Yaskawa INFORM job: -DEFRO-70_PRZYLACZE_60_STARE.JBI

/JOB
//NAME -DEFRO-70_PRZYLACZE_60_STARE
//POS
///NPOS 165,165,165,0,0,0
///TOOL 0
///POSTYPE PULSE
///PULSE
C00000=-281,-101163,-84214,3730,-80188,-1936
C00001=-283,-101162,-84213,3710,-80188,-1936
C00002=115939,-17843,-44700,-6904,-63515,59085
C00003=117854,12047,-44285,-6364,-54274,83125
C00004=118072,11991,-44277,-6360,-54292,83048
C00005=124625,19348,-37580,2226,-58698,65873
C00006=128138,4548,-53928,8815,-39472,48638
C00007=140958,30570,-37086,38951,-57450,21007
C00008=144303,30296,-42198,53003,-55772,9063
C00009=140286,42517,-25172,35381,-64941,20617
C00010=134888,48773,-14255,24473,-68176,15010
C00011=126216,57142,-1405,12520,-73831,-5965
C00012=119431,58070,-113,1607,-75333,-12308
C00013=112362,60124,-1581,-7248,-81906,-32507
C00014=102321,53890,-14377,-28322,-78386,-34401
C00015=102712,42577,-23807,-28139,-73777,-45229
C00016=111795,28445,-30470,-11492,-65646,-58750
C00017=113823,16078,-41175,-14074,-58178,-74794
C00018=114023,15964,-41317,-14088,-58122,-74856
C00019=114170,-2374,-36949,-11645,-74681,-76938
C00020=113314,-7643,-38017,-11019,-76954,88145
C00021=103795,24169,-32802,-5113,-62316,87115
C00022=105717,22963,-33847,-2915,-61383,82248
C00023=105949,12675,-44086,-6804,-51663,75716
C00024=112305,4286,-54083,4280,-38458,55374
C00025=119011,7063,-54209,24198,-38298,40510
C00026=126176,29519,-37310,40709,-52379,12824
C00027=124287,36853,-27992,32882,-57796,17661
C00028=118323,57808,-3223,17808,-73635,15605
C00029=113918,55938,-2510,14235,-71141,-2239
C00030=100452,57135,-1831,-9316,-72769,-11707
C00031=101122,66320,5615,-3405,-83775,-29323
C00032=90969,64062,-2652,-23907,-83052,-31977
C00033=91048,41774,-22566,-24453,-68601,-40164
C00034=95890,27642,-32117,-16170,-61880,-54638
C00035=99625,19836,-37924,-13704,-58629,-70011
C00036=99745,19765,-37997,-13694,-58605,-70048
C00037=99303,8604,-31154,-10952,-72489,-71699
C00038=89422,16015,-23794,-2157,-75183,91094
C00039=91342,36521,-20369,-2557,-66713,90648
C00040=96608,27573,-29625,3606,-58513,75053
C00041=104075,24092,-36197,17400,-51418,55933
C00042=113942,24510,-45627,50308,-45587,24643
C00043=113180,34271,-33600,43117,-51129,17495
C00044=105987,58297,-1625,19620,-69218,16598
C00045=102657,59844,2089,16796,-69099,938
C00046=91593,70320,13088,-1311,-78194,-10490
C00047=88532,80640,21579,-3911,-88822,-24498
C00048=80672,78287,14638,-19772,-88445,-29832
C00049=78449,68959,3821,-24282,-82660,-32911
C00050=77699,46922,-17540,-28065,-68732,-40538
C00051=80754,29721,-31897,-24408,-56253,-47712
C00052=85616,26363,-32270,-14653,-55936,-57384
C00053=85063,22114,-18753,-9149,-74798,-67250
C00054=72786,31521,-9549,-9445,-75352,93043
C00055=79344,46650,-9742,-3090,-64918,94922
C00056=79851,45963,-10489,-3142,-64795,94764
C00057=83555,34866,-22970,1140,-53515,77559
C00058=88637,21070,-41506,13142,-33787,59480
C00059=92546,17739,-49130,33624,-25291,42497
C00060=100296,32921,-36962,50214,-42105,29169
C00061=99518,40044,-26222,41163,-46688,21660
C00062=98807,50157,-13852,39808,-52940,6845
C00063=91319,71721,15887,17155,-70404,4779
C00064=77791,87178,32687,-9256,-82589,-4510
C00065=78950,98816,44020,-1274,-94156,-21475
C00066=71782,98188,39845,-16228,-95193,-28058
C00067=67733,74026,11935,-24954,-78838,-32081
C00068=70123,56840,-3457,-20485,-67729,-42469
C00069=71488,56179,-3109,-17368,-68202,-45369
C00070=72709,50202,-8538,-17621,-67542,-57502
C00071=75039,37514,-3449,-7701,-77257,-64173
C00072=74616,28156,-12897,-9694,-74827,92488
C00073=75521,47327,-9742,-11513,-65249,93468
C00074=83421,34104,-23568,1133,-53536,80045
C00075=88561,20457,-41927,13093,-33823,59529
C00076=92662,18115,-48904,33764,-25272,42413
C00077=97937,26210,-42655,47625,-35211,32454
C00078=99376,40032,-26365,41218,-46566,21666
C00079=100200,49079,-17087,46041,-52311,4065
C00080=91093,71344,15665,17037,-69989,4842
C00081=77993,87860,33884,-9296,-82933,-4594
C00082=79105,99458,45109,-1336,-94484,-21522
C00083=71734,96974,38291,-16203,-94882,-27999
C00084=67577,72994,10856,-25287,-78095,-32283
C00085=72681,51483,-6944,-14654,-65784,-51471
C00086=76109,49503,-7560,-9343,-66865,-57435
C00087=74844,35432,-1015,-7610,-79822,-64270
C00088=74616,28156,-12897,-9694,-74827,92488
C00089=90411,-2677,-20047,-11125,-84138,86440
C00090=90413,-2674,-20051,-11105,-84138,86441
C00091=137757,-12075,-30464,2646,-72394,74401
C00092=139263,-65150,-85436,14259,-28990,73053
C00093=136879,-25803,-69250,35998,-11820,63023
C00094=139290,-23505,-65815,37849,-15870,40588
C00095=138255,-25667,-68923,45072,-10125,18948
C00096=137540,-11621,-49291,15825,-29065,282
C00097=134494,-8817,-45605,4069,-31945,-3289
C00098=134604,-8591,-45393,4272,-32069,-3452
C00099=128608,-126,-37091,-12913,-41572,-17604
C00100=135365,-22598,-63276,22384,-16411,-55250
C00101=133643,-21758,-61840,7774,-18256,-58833
C00102=132849,-22230,-62300,-146,-18489,-67744
C00103=134650,-26769,-71812,22381,-6082,-94556
C00104=132637,-74135,-100376,4983,-10333,-85647
C00105=119687,-78067,-87939,-2788,-20735,84624
C00106=119992,-27745,-68017,-3051,-15116,84333
C00107=119030,-28696,-69591,-21999,-13157,75803
C00108=119146,-27568,-67331,-20983,-14326,49763
C00109=119106,-25320,-64288,-16073,-16150,28459
C00110=116990,-27787,-67992,-36968,-13306,28443
C00111=114451,-20387,-59191,-34974,-24024,21051
C00112=114289,-23226,-63137,-42813,-20195,20855
C00113=115755,-27101,-67787,-45506,-13897,17108
C00114=116631,-28534,-69574,-43897,-10967,13052
C00115=119721,-30747,-72526,-5019,-4908,-12317
C00116=124673,-29524,-70968,54153,-12690,-50315
C00117=110381,-14519,-53439,-34713,-36084,-50985
C00118=115065,-20808,-58231,-19385,-28009,-64203
C00119=113126,-78683,-102705,-45607,-16425,-60367
C00120=120908,-77676,-80309,7462,-22023,84016
C00121=119355,-30092,-72700,-7480,-8883,86833
C00122=119330,-30666,-73900,-37441,-7256,75668
C00123=119392,-31005,-74194,-36731,-7285,75171
C00124=119107,-25533,-64139,-15884,-16345,28370
C00125=118189,-11113,-47154,-8478,-33276,7215
C00126=118285,-13415,-49709,-5227,-31034,-7778
C00127=112204,-14619,-53166,-28572,-30616,-12922
C00128=112459,-20642,-60567,-34495,-24493,-27463
C00129=113253,-23242,-63602,-34662,-21946,-37788
C00130=117822,-27208,-67860,-16762,-15410,-62087
C00131=114088,-29625,-74008,-62760,-13130,-51071
C00132=113074,-79856,-103225,-44998,-16651,-60643
C00133=120443,-70015,-86553,-1670,-18639,84017
C00134=119855,-29453,-70963,-4444,-11447,85360
C00135=119350,-27114,-66909,-10824,-16764,76179
C00136=120538,-28712,-69581,-9042,-12118,60389
C00137=121453,-23804,-62042,-1822,-20367,42740
C00138=119104,-25714,-64462,-15988,-16245,28420
C00139=118127,-25090,-63854,-17709,-16479,10287
C00140=118054,-20647,-58029,-8598,-22594,-6818
C00141=116391,-17852,-55102,-12391,-26715,-16410
C00142=113676,-17333,-55635,-24105,-28107,-26621
C00143=114148,-20487,-59353,-25400,-25301,-39443
C00144=114654,-26064,-67349,-36235,-17702,-47147
C00145=115014,-30497,-76060,-73901,-10838,-47744
C00146=112648,-89264,-107216,-40476,-18619,-62704
C00147=115490,-77010,-93554,-11224,-18305,89052
C00148=125433,-24819,-64014,25600,-22035,67229
C00149=124409,-21324,-58576,14136,-26697,62401
C00150=126029,-28427,-71429,47699,-12406,35561
C00151=126376,-14543,-51553,17453,-33391,37954
C00152=119104,-25707,-64456,-15987,-16243,28419
C00153=102227,-21803,-62565,-47260,-20333,28942
C00154=103256,-22698,-63333,-30550,-15064,8897
C00155=100032,-11798,-50575,-26640,-29993,-6479
C00156=97406,-10335,-50320,-35130,-33056,-18084
C00157=102127,-19671,-59474,-25169,-24074,-49644
C00158=96594,-22492,-70681,-79494,-21703,-41695
C00159=112538,-91654,-108181,-39431,-19159,-63177
C00160=113545,-73371,-70378,-16072,-42358,69017
C00161=89593,-90202,-78264,-12204,-55560,23671
C00162=60247,-88344,-77535,-12630,-64499,59028
C00163=11932,-100155,-87763,417,-74819,10359
C00164=-281,-101163,-84214,3730,-80188,-1936
BC00000=570125
BC00001=868704
BC00002=878894
BC00003=878037
BC00004=878037
BC00005=878038
BC00006=878037
BC00007=878038
BC00008=878038
BC00009=878038
BC00010=878038
BC00011=878038
BC00012=878038
BC00013=878037
BC00014=878037
BC00015=878037
BC00016=878037
BC00017=878037
BC00018=878037
BC00019=878037
BC00020=912823
BC00021=878035
BC00022=878036
BC00023=878036
BC00024=878037
BC00025=878037
BC00026=878037
BC00027=878037
BC00028=878038
BC00029=878038
BC00030=878037
BC00031=878037
BC00032=878037
BC00033=878037
BC00034=878037
BC00035=878037
BC00036=878037
BC00037=878037
BC00038=878035
BC00039=878036
BC00040=878037
BC00041=878037
BC00042=878038
BC00043=878038
BC00044=878038
BC00045=878038
BC00046=878037
BC00047=878037
BC00048=878037
BC00049=878037
BC00050=878037
BC00051=878037
BC00052=878037
BC00053=878037
BC00054=878037
BC00055=878035
BC00056=878035
BC00057=877203
BC00058=877947
BC00059=878201
BC00060=878342
BC00061=878784
BC00062=877961
BC00063=877604
BC00064=878504
BC00065=878840
BC00066=878535
BC00067=877975
BC00068=879348
BC00069=879174
BC00070=879174
BC00071=878037
BC00072=915550
BC00073=913919
BC00074=916409
BC00075=916569
BC00076=916479
BC00077=916387
BC00078=916586
BC00079=915550
BC00080=915870
BC00081=916359
BC00082=916889
BC00083=917058
BC00084=916344
BC00085=916664
BC00086=916387
BC00087=915811
BC00088=915550
BC00089=915550
BC00090=915550
BC00091=915550
BC00092=915550
BC00093=915550
BC00094=915550
BC00095=915550
BC00096=915550
BC00097=915550
BC00098=915550
BC00099=915550
BC00100=915550
BC00101=915550
BC00102=915550
BC00103=915550
BC00104=915550
BC00105=915550
BC00106=915551
BC00107=915550
BC00108=915550
BC00109=915550
BC00110=915550
BC00111=915550
BC00112=915550
BC00113=915550
BC00114=915550
BC00115=915550
BC00116=915550
BC00117=915550
BC00118=915550
BC00119=915550
BC00120=954211
BC00121=953187
BC00122=954162
BC00123=954160
BC00124=954071
BC00125=953684
BC00126=953455
BC00127=953244
BC00128=953665
BC00129=953702
BC00130=953799
BC00131=953749
BC00132=953683
BC00133=992214
BC00134=992214
BC00135=992103
BC00136=991968
BC00137=992423
BC00138=992186
BC00139=992082
BC00140=991590
BC00141=991168
BC00142=991569
BC00143=992150
BC00144=992735
BC00145=991845
BC00146=991844
BC00147=1026906
BC00148=1030289
BC00149=1030277
BC00150=1030261
BC00151=1030281
BC00152=1030485
BC00153=997557
BC00154=991657
BC00155=991168
BC00156=991569
BC00157=992735
BC00158=991845
BC00159=1030552
BC00160=1030552
BC00161=1015004
BC00162=995119
BC00163=847363
BC00164=570125
EC00000=1163,0
EC00001=1166,0
EC00002=-1742,0
EC00003=-1741,0
EC00004=-1741,0
EC00005=-1743,0
EC00006=-1742,0
EC00007=-1741,0
EC00008=-1741,0
EC00009=-1741,0
EC00010=-1741,0
EC00011=-1741,0
EC00012=-1741,0
EC00013=-1741,0
EC00014=-1742,0
EC00015=-1742,0
EC00016=-1742,0
EC00017=-1741,0
EC00018=-1741,0
EC00019=-1741,0
EC00020=-1741,0
EC00021=-1745,0
EC00022=-1744,0
EC00023=-1743,0
EC00024=-1742,0
EC00025=-1742,0
EC00026=-1741,0
EC00027=-1741,0
EC00028=-1741,0
EC00029=-1741,0
EC00030=-1741,0
EC00031=-1741,0
EC00032=-1742,0
EC00033=-1742,0
EC00034=-1741,0
EC00035=-1741,0
EC00036=-1741,0
EC00037=-1741,0
EC00038=-1743,0
EC00039=-1742,0
EC00040=-1742,0
EC00041=-1742,0
EC00042=-1741,0
EC00043=-1741,0
EC00044=-1595,0
EC00045=-1742,0
EC00046=-1741,0
EC00047=-1741,0
EC00048=-1742,0
EC00049=-1742,0
EC00050=-1742,0
EC00051=-1742,0
EC00052=-1742,0
EC00053=-1741,0
EC00054=-1741,0
EC00055=-1743,0
EC00056=-1743,0
EC00057=-1742,0
EC00058=-1743,0
EC00059=-1742,0
EC00060=-1741,0
EC00061=-1741,0
EC00062=-1742,0
EC00063=-1742,0
EC00064=-1742,0
EC00065=-1741,0
EC00066=-1741,0
EC00067=-1741,0
EC00068=-1741,0
EC00069=-1741,0
EC00070=-1741,0
EC00071=-1741,0
EC00072=-1741,0
EC00073=-1742,0
EC00074=-1742,0
EC00075=-1743,0
EC00076=-1742,0
EC00077=-1741,0
EC00078=-1740,0
EC00079=-1742,0
EC00080=-1742,0
EC00081=-1742,0
EC00082=-1741,0
EC00083=-1741,0
EC00084=-1741,0
EC00085=-1742,0
EC00086=-1742,0
EC00087=-1741,0
EC00088=-1741,0
EC00089=-1741,0
EC00090=-84878,0
EC00091=-84879,0
EC00092=-84877,0
EC00093=-84877,0
EC00094=-84877,0
EC00095=-84877,0
EC00096=-84877,0
EC00097=-84877,0
EC00098=-84877,0
EC00099=-84877,0
EC00100=-84877,0
EC00101=-84877,0
EC00102=-84877,0
EC00103=-84877,0
EC00104=-84877,0
EC00105=-84877,0
EC00106=-84878,0
EC00107=-84877,0
EC00108=-84877,0
EC00109=-84877,0
EC00110=-84877,0
EC00111=-84877,0
EC00112=-84877,0
EC00113=-84877,0
EC00114=-84877,0
EC00115=-84877,0
EC00116=-84877,0
EC00117=-84877,0
EC00118=-84877,0
EC00119=-84877,0
EC00120=-84877,0
EC00121=-84878,0
EC00122=-84877,0
EC00123=-84877,0
EC00124=-84877,0
EC00125=-84877,0
EC00126=-84877,0
EC00127=-84877,0
EC00128=-84877,0
EC00129=-84877,0
EC00130=-84877,0
EC00131=-84877,0
EC00132=-84877,0
EC00133=-84877,0
EC00134=-84877,0
EC00135=-84877,0
EC00136=-84877,0
EC00137=-84877,0
EC00138=-84877,0
EC00139=-84877,0
EC00140=-84877,0
EC00141=-84877,0
EC00142=-84877,0
EC00143=-84877,0
EC00144=-84877,0
EC00145=-84877,0
EC00146=-84877,0
EC00147=-84877,0
EC00148=-84877,0
EC00149=-84877,0
EC00150=-84877,0
EC00151=-84877,0
EC00152=-84877,0
EC00153=-84877,0
EC00154=-84877,0
EC00155=-84877,0
EC00156=-84877,0
EC00157=-84877,0
EC00158=-84877,0
EC00159=-84877,0
EC00160=-84877,0
EC00161=-1879,0
EC00162=-1342,0
EC00163=498,0
EC00164=1163,0
//INST
///DATE 2025/05/12 13:13
///COMM OZZ
///ATTR SC,RW
///GROUP1 RB1,BS1
///GROUP2 ST1
NOP
MOVJ C00000 BC00000 VJ=70.00 DEC=20  +MOVJ EC00000 VJ=70.00
MOVJ C00001 BC00001 VJ=40.00 DEC=20  +MOVJ EC00001 VJ=40.00
MOVJ C00002 BC00002 VJ=70.00 DEC=20  +MOVJ EC00002 VJ=70.00
MOVJ C00003 BC00003 VJ=40.00 DEC=20  +MOVJ EC00003 VJ=70.00
MACRO1 MJ#(0) ARGF8
WVON WEV#(1)
ARCON
MOVC C00004 BC00004 V=4.2 DEC=20  +MOVJ EC00004 VJ=70.00
MOVC C00005 BC00005 V=4.2 DEC=20  +MOVJ EC00005 VJ=30.00
MOVC C00006 BC00006 V=4.2 DEC=20  +MOVJ EC00006 VJ=30.00
MOVC C00007 BC00007 V=4.2 DEC=20  +MOVJ EC00007 VJ=30.00
MOVC C00008 BC00008 V=4.2 DEC=20  +MOVJ EC00008 VJ=30.00
MOVC C00009 BC00009 V=4.2 DEC=20  +MOVJ EC00009 VJ=0.78
MOVC C00010 BC00010 V=4.2 DEC=20  +MOVJ EC00010 VJ=30.00
MOVC C00011 BC00011 V=4.2 DEC=20  +MOVJ EC00011 VJ=30.00
MOVC C00012 BC00012 V=4.2 DEC=20  +MOVJ EC00012 VJ=30.00
MOVC C00013 BC00013 V=4.2 DEC=20  +MOVJ EC00013 VJ=30.00
MOVC C00014 BC00014 V=4.2 DEC=20  +MOVJ EC00014 VJ=30.00
MOVC C00015 BC00015 V=4.2 DEC=20  +MOVJ EC00015 VJ=30.00
MOVC C00016 BC00016 V=4.2 DEC=20  +MOVJ EC00016 VJ=30.00
MOVC C00017 BC00017 V=4.2 DEC=20  +MOVJ EC00017 VJ=30.00
MOVJ C00018 BC00018 VJ=30.00 DEC=20  +MOVJ EC00018 VJ=30.00
WVOF
ARCOF
MOVJ C00019 BC00019 VJ=40.00 DEC=20  +MOVJ EC00019 VJ=40.00
MOVJ C00020 BC00020 VJ=70.00 DEC=20  +MOVJ EC00020 VJ=0.78
MOVJ C00021 BC00021 VJ=30.00 DEC=20  +MOVJ EC00021 VJ=0.78
MACRO1 MJ#(0) ARGF8
WVON WEV#(1)
ARCON
MOVC C00022 BC00022 V=4.2 DEC=20  +MOVJ EC00022 VJ=0.78
MOVC C00023 BC00023 V=4.2 DEC=20  +MOVJ EC00023 VJ=0.78
MOVC C00024 BC00024 V=4.2 DEC=20  +MOVJ EC00024 VJ=30.00
MOVC C00025 BC00025 V=4.2 DEC=20  +MOVJ EC00025 VJ=30.00
MOVC C00026 BC00026 V=5.0 DEC=20  +MOVJ EC00026 VJ=30.00
MOVC C00027 BC00027 V=4.2 DEC=20  +MOVJ EC00027 VJ=0.78
MOVC C00028 BC00028 V=4.2 DEC=20  +MOVJ EC00028 VJ=30.00
MOVC C00029 BC00029 V=4.2 DEC=20  +MOVJ EC00029 VJ=30.00
MOVC C00030 BC00030 V=4.2 DEC=20  +MOVJ EC00030 VJ=30.00
MOVC C00031 BC00031 V=4.2 DEC=20  +MOVJ EC00031 VJ=30.00
MOVC C00032 BC00032 V=4.2 DEC=20  +MOVJ EC00032 VJ=30.00
MOVC C00033 BC00033 V=4.2 DEC=20  +MOVJ EC00033 VJ=30.00
MOVC C00034 BC00034 V=4.2 DEC=20  +MOVJ EC00034 VJ=30.00
MOVC C00035 BC00035 V=4.2 DEC=20  +MOVJ EC00035 VJ=30.00
MOVJ C00036 BC00036 VJ=25.00 DEC=20  +MOVJ EC00036 VJ=30.00
WVOF
ARCOF
MOVJ C00037 BC00037 VJ=30.00 DEC=20  +MOVJ EC00037 VJ=30.00
MOVJ C00038 BC00038 VJ=30.00 DEC=20  +MOVJ EC00038 VJ=30.00
MOVJ C00039 BC00039 VJ=30.00 DEC=20  +MOVJ EC00039 VJ=30.00
WVON WEV#(1)
ARCON
MOVC C00040 BC00040 V=4.2 DEC=20  +MOVJ EC00040 VJ=30.00
MOVC C00041 BC00041 V=4.2 DEC=20  +MOVJ EC00041 VJ=30.00
MOVC C00042 BC00042 V=4.2 DEC=20  +MOVJ EC00042 VJ=30.00
MOVC C00043 BC00043 V=4.2 DEC=20  +MOVJ EC00043 VJ=30.00
MOVC C00044 BC00044 V=4.2 DEC=20  +MOVJ EC00044 VJ=30.00
MOVC C00045 BC00045 V=4.2 DEC=20  +MOVJ EC00045 VJ=30.00
MOVC C00046 BC00046 V=4.2 DEC=20  +MOVJ EC00046 VJ=30.00
MOVC C00047 BC00047 V=4.2 DEC=20  +MOVJ EC00047 VJ=30.00
MOVC C00048 BC00048 V=4.2 DEC=20  +MOVJ EC00048 VJ=30.00
MOVC C00049 BC00049 V=4.2 DEC=20  +MOVJ EC00049 VJ=0.78
MOVC C00050 BC00050 V=5.8 DEC=20  +MOVJ EC00050 VJ=30.00
MOVC C00051 BC00051 V=4.2 DEC=20  +MOVJ EC00051 VJ=0.78
MOVC C00052 BC00052 V=4.2 DEC=20  +MOVJ EC00052 VJ=30.00
ARCOF
WVOF
MOVJ C00053 BC00053 VJ=30.00 DEC=20  +MOVJ EC00053 VJ=30.00
MOVJ C00054 BC00054 VJ=30.00 DEC=20  +MOVJ EC00054 VJ=30.00
MOVJ C00055 BC00055 VJ=30.00 DEC=20  +MOVJ EC00055 VJ=30.00
WVON WEV#(1)
ARCON
MOVC C00056 BC00056 V=4.2 DEC=20  +MOVJ EC00056 VJ=0.78
MOVC C00057 BC00057 V=4.2 DEC=20  +MOVJ EC00057 VJ=0.78
MOVC C00058 BC00058 V=4.2 DEC=20  +MOVJ EC00058 VJ=0.78
MOVC C00059 BC00059 V=4.2 DEC=20  +MOVJ EC00059 VJ=0.78
MOVC C00060 BC00060 V=4.2 DEC=20  +MOVJ EC00060 VJ=0.78
MOVC C00061 BC00061 V=4.2 DEC=20  +MOVJ EC00061 VJ=0.78
MOVC C00062 BC00062 V=4.2 DEC=20  +MOVJ EC00062 VJ=0.78
MOVC C00063 BC00063 V=4.2 DEC=20  +MOVJ EC00063 VJ=0.78
MOVC C00064 BC00064 V=4.2 DEC=20  +MOVJ EC00064 VJ=0.78
MOVC C00065 BC00065 V=4.2 DEC=20  +MOVJ EC00065 VJ=0.78
MOVC C00066 BC00066 V=4.2 DEC=20  +MOVJ EC00066 VJ=0.78
MOVC C00067 BC00067 V=4.2 DEC=20  +MOVJ EC00067 VJ=0.78
MOVC C00068 BC00068 V=4.2 DEC=20  +MOVJ EC00068 VJ=0.78
MOVC C00069 BC00069 V=4.2 DEC=20  +MOVJ EC00069 VJ=0.78
MOVC C00070 BC00070 V=4.2 DEC=20  +MOVJ EC00070 VJ=0.78
WVOF
ARCOF
MOVJ C00071 BC00071 VJ=30.00 DEC=20  +MOVJ EC00071 VJ=30.00
MOVJ C00072 BC00072 VJ=30.00 DEC=20  +MOVJ EC00072 VJ=30.00
MOVJ C00073 BC00073 VJ=30.00 DEC=20  +MOVJ EC00073 VJ=30.00
WVON WEV#(1)
ARCON
MOVC C00074 BC00074 V=4.2 DEC=20  +MOVJ EC00074 VJ=30.00
MOVC C00075 BC00075 V=4.2 DEC=20  +MOVJ EC00075 VJ=30.00
MOVC C00076 BC00076 V=4.2 DEC=20  +MOVJ EC00076 VJ=40.00
MOVC C00077 BC00077 V=4.2 DEC=20  +MOVJ EC00077 VJ=30.00
MOVC C00078 BC00078 V=4.2 DEC=20  +MOVJ EC00078 VJ=25.00
MOVC C00079 BC00079 V=4.2 DEC=20  +MOVJ EC00079 VJ=30.00
MOVC C00080 BC00080 V=4.2 DEC=20  +MOVJ EC00080 VJ=70.00
MOVC C00081 BC00081 V=4.2 DEC=20  +MOVJ EC00081 VJ=30.00
MOVC C00082 BC00082 V=4.2 DEC=20  +MOVJ EC00082 VJ=30.00
MOVC C00083 BC00083 V=4.2 DEC=20  +MOVJ EC00083 VJ=30.00
MOVC C00084 BC00084 V=4.2 DEC=20  +MOVJ EC00084 VJ=30.00
MOVC C00085 BC00085 V=4.2 DEC=20  +MOVJ EC00085 VJ=0.78
MOVC C00086 BC00086 V=4.2 DEC=20  +MOVJ EC00086 VJ=30.00
ARCOF
WVOF
MOVJ C00087 BC00087 VJ=30.00 DEC=20  +MOVJ EC00087 VJ=30.00
MOVJ C00088 BC00088 VJ=30.00 DEC=20  +MOVJ EC00088 VJ=30.00
MOVJ C00089 BC00089 VJ=30.00 DEC=20  +MOVJ EC00089 VJ=30.00
MOVJ C00090 BC00090 VJ=30.00 DEC=20  +MOVJ EC00090 VJ=30.00
MOVJ C00091 BC00091 VJ=30.00 DEC=20  +MOVJ EC00091 VJ=30.00
MOVJ C00092 BC00092 VJ=70.00 DEC=20  +MOVJ EC00092 VJ=0.78
MOVJ C00093 BC00093 VJ=30.00 DEC=20  +MOVJ EC00093 VJ=0.78
MACRO1 MJ#(0) ARGF4
ARCON
MOVC C00094 BC00094 V=5.0 DEC=20  +MOVJ EC00094 VJ=0.78
MOVC C00095 BC00095 V=5.0 DEC=20  +MOVJ EC00095 VJ=0.78
MOVC C00096 BC00096 V=5.0 DEC=20  +MOVJ EC00096 VJ=0.78
MOVC C00097 BC00097 V=5.0 DEC=20  +MOVJ EC00097 VJ=0.78
MOVC C00098 BC00098 V=5.0 DEC=20  +MOVJ EC00098 VJ=0.78
MOVC C00099 BC00099 V=5.0 DEC=20  +MOVJ EC00099 VJ=0.78
MOVC C00100 BC00100 V=5.0 DEC=20  +MOVJ EC00100 VJ=0.78
MOVC C00101 BC00101 V=5.0 DEC=20  +MOVJ EC00101 VJ=0.78
MOVC C00102 BC00102 V=5.0 DEC=20  +MOVJ EC00102 VJ=0.78
MOVC C00103 BC00103 V=5.0 DEC=20  +MOVJ EC00103 VJ=0.78
ARCOF
MOVJ C00104 BC00104 VJ=40.00 DEC=20  +MOVJ EC00104 VJ=0.78
MOVJ C00105 BC00105 VJ=40.00 DEC=20  +MOVJ EC00105 VJ=0.78
MOVJ C00106 BC00106 VJ=40.00 DEC=20  +MOVJ EC00106 VJ=0.78
ARCON
MOVC C00107 BC00107 V=5.0 DEC=20  +MOVJ EC00107 VJ=0.78
MOVC C00108 BC00108 V=5.0 DEC=20  +MOVJ EC00108 VJ=40.00
MOVC C00109 BC00109 V=5.0 DEC=20  +MOVJ EC00109 VJ=0.78
MOVC C00110 BC00110 V=5.0 DEC=20  +MOVJ EC00110 VJ=0.78
MOVC C00111 BC00111 V=5.0 DEC=20  +MOVJ EC00111 VJ=0.78
MOVC C00112 BC00112 V=5.0 DEC=20  +MOVJ EC00112 VJ=0.78
MOVL C00113 BC00113 V=5.0 DEC=20  +MOVJ EC00113 VJ=80.00
MOVC C00114 BC00114 V=5.0 DEC=20  +MOVJ EC00114 VJ=0.78
MOVC C00115 BC00115 V=5.0 DEC=20  +MOVJ EC00115 VJ=0.78
MOVC C00116 BC00116 V=5.0 DEC=20  +MOVJ EC00116 VJ=0.78
MOVC C00117 BC00117 V=5.0 DEC=20  +MOVJ EC00117 VJ=70.00
MOVC C00118 BC00118 V=5.0 DEC=20  +MOVJ EC00118 VJ=0.78
ARCOF
MOVJ C00119 BC00119 VJ=40.00 DEC=20  +MOVJ EC00119 VJ=0.78
MOVJ C00120 BC00120 VJ=40.00 DEC=20  +MOVJ EC00120 VJ=0.78
MOVJ C00121 BC00121 VJ=40.00 DEC=20  +MOVJ EC00121 VJ=0.78
ARCON
MOVC C00122 BC00122 V=5.0 DEC=20  +MOVJ EC00122 VJ=0.78
MOVC C00123 BC00123 V=5.0 DEC=20  +MOVJ EC00123 VJ=0.78
MOVC C00124 BC00124 V=5.0 DEC=20  +MOVJ EC00124 VJ=0.78
MOVC C00125 BC00125 V=5.0 DEC=20  +MOVJ EC00125 VJ=0.78
MOVC C00126 BC00126 V=5.0 DEC=20  +MOVJ EC00126 VJ=0.78
MOVC C00127 BC00127 V=5.0 DEC=20  +MOVJ EC00127 VJ=0.78
MOVC C00128 BC00128 V=5.0 DEC=20  +MOVJ EC00128 VJ=0.78
MOVC C00129 BC00129 V=5.0 DEC=20  +MOVJ EC00129 VJ=0.78
MOVC C00130 BC00130 V=5.0 DEC=20  +MOVJ EC00130 VJ=0.78
MOVC C00131 BC00131 V=5.0 DEC=20  +MOVJ EC00131 VJ=0.78
ARCOF
MOVJ C00132 BC00132 VJ=40.00 DEC=20  +MOVJ EC00132 VJ=0.78
MOVJ C00133 BC00133 VJ=40.00 DEC=20  +MOVJ EC00133 VJ=0.78
MOVJ C00134 BC00134 VJ=40.00 DEC=20  +MOVJ EC00134 VJ=0.78
ARCON
MOVC C00135 BC00135 V=5.0 DEC=20  +MOVJ EC00135 VJ=0.78
MOVC C00136 BC00136 V=5.0 DEC=20  +MOVJ EC00136 VJ=0.78
MOVC C00137 BC00137 V=5.0 DEC=20  +MOVJ EC00137 VJ=0.78
MOVC C00138 BC00138 V=5.0 DEC=20  +MOVJ EC00138 VJ=0.78
MOVC C00139 BC00139 V=5.0 DEC=20  +MOVJ EC00139 VJ=0.78
MOVC C00140 BC00140 V=5.0 DEC=20  +MOVJ EC00140 VJ=0.78
MOVC C00141 BC00141 V=5.0 DEC=20  +MOVJ EC00141 VJ=0.78
MOVC C00142 BC00142 V=5.0 DEC=20  +MOVJ EC00142 VJ=0.78
MOVC C00143 BC00143 V=5.0 DEC=20  +MOVJ EC00143 VJ=0.78
MOVC C00144 BC00144 V=5.0 DEC=20  +MOVJ EC00144 VJ=0.78
MOVC C00145 BC00145 V=5.0 DEC=20  +MOVJ EC00145 VJ=0.78
ARCOF
MOVJ C00146 BC00146 VJ=40.00 DEC=20  +MOVJ EC00146 VJ=0.78
MOVJ C00147 BC00147 VJ=40.00 DEC=20  +MOVJ EC00147 VJ=0.78
MOVJ C00148 BC00148 VJ=40.00 DEC=20  +MOVJ EC00148 VJ=0.78
ARCON
MOVC C00149 BC00149 V=5.0 DEC=20  +MOVJ EC00149 VJ=0.78
MOVC C00150 BC00150 V=5.0 DEC=20  +MOVJ EC00150 VJ=0.78
MOVC C00151 BC00151 V=5.0 DEC=20  +MOVJ EC00151 VJ=0.78
MOVC C00152 BC00152 V=5.0 DEC=20  +MOVJ EC00152 VJ=0.78
MOVC C00153 BC00153 V=5.0 DEC=20  +MOVJ EC00153 VJ=70.00
MOVC C00154 BC00154 V=5.0 DEC=20  +MOVJ EC00154 VJ=30.00
MOVC C00155 BC00155 V=5.0 DEC=20  +MOVJ EC00155 VJ=70.00
MOVC C00156 BC00156 V=5.0 DEC=20  +MOVJ EC00156 VJ=70.00
MOVC C00157 BC00157 V=5.0 DEC=20  +MOVJ EC00157 VJ=70.00
MOVC C00158 BC00158 V=5.0 DEC=20  +MOVJ EC00158 VJ=70.00
ARCOF
MOVJ C00159 BC00159 VJ=40.00 DEC=20  +MOVJ EC00159 VJ=0.78
MOVJ C00160 BC00160 VJ=40.00 DEC=20  +MOVJ EC00160 VJ=0.78
MOVJ C00161 BC00161 VJ=40.00 DEC=20  +MOVJ EC00161 VJ=40.00
MOVJ C00162 BC00162 VJ=70.00 DEC=20  +MOVJ EC00162 VJ=0.78
MOVJ C00163 BC00163 VJ=70.00 DEC=20  +MOVJ EC00163 VJ=70.00
MOVJ C00164 BC00164 VJ=40.00 DEC=20  +MOVJ EC00164 VJ=0.78
END
